(* IEC 61131-3 sources: SemaPLC/sema-plc-benchmark/spec2control-benchmark/data/st-baseline/desalination/pous/programs, 6 files *)

(* ---- main.st ---- *)
PROGRAM main
VAR
	Heartbeat : bool;
END_VAR

(* Entry point required by OpenPLC Editor v4. The process sections run as parallel program instances under task0; main only provides a scan heartbeat. *)
Heartbeat := NOT Heartbeat;

END_PROGRAM

(* ---- Section2.st ---- *)
PROGRAM Section2
VAR
	FT101_Flow_PV : real;
	FT102_Flow_PV : real;
	AT101_Analyzer_PV : real;
	AT103_Analyzer_PV : real;
	LT104_Level_PV : real;
	LT105_Level_PV : real;
	FC101_MV_Out : real;
	FC102_MV_Out : real;
	FV101_Valve_Position : real;
	FV102_Valve_Position : real;
	SP101_PctCmd : real;
	SP102_PctCmd : real;
	FlowDevAlarm101 : bool;
	FlowDevAlarm102 : bool;
	AT_101 : ANALOG_IN;
	AT_103 : ANALOG_IN;
	FC_101 : PID_BASIC;
	FC_102 : PID_BASIC;
	FT_101 : ANALOG_IN;
	FT_102 : ANALOG_IN;
	FV_101 : VALVE_ELECTRIC;
	FV_102 : VALVE_ELECTRIC;
	LT_104 : ANALOG_IN;
	LT_105 : ANALOG_IN;
	XV_102 : VALVE_ON_OFF;
	SP101_DevDelay_TON : TON;
	SP102_DevDelay_TON : TON;
	XV102NotOpen_NOT : bool;
	Contamination_OR : bool;
	FV101_Inhibit_OR : bool;
	FV102_Inhibit_OR : bool;
	SP101_PctNorm_DIV : real;
	SP101_PctScaled_MULT : real;
	SP101_PctOffset_ADD : real;
	SP101_PctToFrac_DIV : real;
	SP101_SP_EU_MULT : real;
	DL101_MULT : real;
	SP101_1p1_MULT : real;
	SP101_0p9_MULT : real;
	SP101_PV_GT_HighThresh : bool;
	SP101_PV_LT_LowThresh : bool;
	SP101_DevBand_OR : bool;
	SP102_PctNorm_DIV : real;
	SP102_PctScaled_MULT : real;
	SP102_PctOffset_ADD : real;
	SP102_PctToFrac_DIV : real;
	SP102_SP_EU_MULT : real;
	DL102_MULT : real;
	SP102_1p1_MULT : real;
	SP102_0p9_MULT : real;
	SP102_PV_GT_HighThresh : bool;
	SP102_PV_LT_LowThresh : bool;
	SP102_DevBand_OR : bool;
END_VAR

AT_101(
    PV_High := 50.0,
    Alarm_Enable := TRUE);
AT_103(
    PV_High := 35.0,
    Alarm_Enable := TRUE);
SP101_PctNorm_DIV := SP101_PctCmd / 100.0;
SP101_PctScaled_MULT := SP101_PctNorm_DIV * 59.0;
SP101_PctOffset_ADD := SP101_PctScaled_MULT + 16.0;
SP101_PctToFrac_DIV := SP101_PctOffset_ADD / 100.0;
SP101_SP_EU_MULT := SP101_PctToFrac_DIV * 5000.0;
DL101_MULT := SP101_SP_EU_MULT * 0.1;
FT_101(
    PV_High := 5500.0,
    PV_Low := 450.0,
    Scaling_Slope := 312.5,
    Scaling_Offset := -1250.0,
    Alarm_Enable := TRUE);
FC_101(
    AUTO := TRUE,
    PV := FT_101.PV,
    SP := SP101_SP_EU_MULT,
    MV_MIN := 0.0,
    MV_MAX := 100.0,
    X0 := 0.0,
    KP := 2.5,
    TR := 0.8,
    TD := 0.2,
    Deviation_Limit := DL101_MULT,
    Inhibit := FT_101.General_Fault);
SP102_PctNorm_DIV := SP102_PctCmd / 100.0;
SP102_PctScaled_MULT := SP102_PctNorm_DIV * 59.0;
SP102_PctOffset_ADD := SP102_PctScaled_MULT + 16.0;
SP102_PctToFrac_DIV := SP102_PctOffset_ADD / 100.0;
SP102_SP_EU_MULT := SP102_PctToFrac_DIV * 3000.0;
DL102_MULT := SP102_SP_EU_MULT * 0.1;
FT_102(
    PV_High := 3300.0,
    PV_Low := 270.0,
    Scaling_Slope := 187.5,
    Scaling_Offset := -750.0,
    Alarm_Enable := TRUE);
FC_102(
    AUTO := TRUE,
    PV := FT_102.PV,
    SP := SP102_SP_EU_MULT,
    MV_MIN := 0.0,
    MV_MAX := 100.0,
    X0 := 0.0,
    KP := 2.5,
    TR := 0.8,
    TD := 0.2,
    Deviation_Limit := DL102_MULT,
    Inhibit := FT_102.General_Fault);
Contamination_OR := AT_101.High_Alarm OR AT_103.High_Alarm;
LT_104(
    PV_Low := 2.0,
    Alarm_Enable := TRUE);
LT_105(
    Alarm_Enable := TRUE);
XV_102(
    Inhibit := Contamination_OR);
XV102NotOpen_NOT := NOT XV_102.FB_Opened;
FV101_Inhibit_OR := XV102NotOpen_NOT OR Contamination_OR OR LT_104.Low_Alarm OR LT_105.High_Alarm OR FT_101.General_Fault;
FV_101(
    Control_Signal := FC_101.XOUT,
    Manual_Mode := FALSE,
    Manual_Position := 0.0,
    Open_Limit := 100.0,
    Close_Limit := 0.0,
    Inhibit := FV101_Inhibit_OR);
FV102_Inhibit_OR := XV102NotOpen_NOT OR Contamination_OR OR LT_104.Low_Alarm OR LT_105.High_Alarm OR FT_102.General_Fault;
FV_102(
    Control_Signal := FC_102.XOUT,
    Manual_Mode := FALSE,
    Manual_Position := 0.0,
    Open_Limit := 100.0,
    Close_Limit := 0.0,
    Inhibit := FV102_Inhibit_OR);
SP101_1p1_MULT := SP101_SP_EU_MULT * 1.1;
SP101_PV_GT_HighThresh := (FT_101.PV > SP101_1p1_MULT);
SP101_0p9_MULT := SP101_SP_EU_MULT * 0.9;
SP101_PV_LT_LowThresh := (FT_101.PV < SP101_0p9_MULT);
SP101_DevBand_OR := SP101_PV_GT_HighThresh OR SP101_PV_LT_LowThresh;
SP101_DevDelay_TON(
    IN := SP101_DevBand_OR,
    PT := T#30s);
SP102_1p1_MULT := SP102_SP_EU_MULT * 1.1;
SP102_PV_GT_HighThresh := (FT_102.PV > SP102_1p1_MULT);
SP102_0p9_MULT := SP102_SP_EU_MULT * 0.9;
SP102_PV_LT_LowThresh := (FT_102.PV < SP102_0p9_MULT);
SP102_DevBand_OR := SP102_PV_GT_HighThresh OR SP102_PV_LT_LowThresh;
SP102_DevDelay_TON(
    IN := SP102_DevBand_OR,
    PT := T#30s);

(* Outputs published to other sections / HMI. *)
FT101_Flow_PV := FT_101.PV;
FT102_Flow_PV := FT_102.PV;
AT101_Analyzer_PV := AT_101.PV;
AT103_Analyzer_PV := AT_103.PV;
LT104_Level_PV := LT_104.PV;
LT105_Level_PV := LT_105.PV;
FC101_MV_Out := FC_101.XOUT;
FC102_MV_Out := FC_102.XOUT;
FV101_Valve_Position := FV_101.Valve_Position;
FV102_Valve_Position := FV_102.Valve_Position;
FlowDevAlarm101 := SP101_DevDelay_TON.Q;
FlowDevAlarm102 := SP102_DevDelay_TON.Q;

END_PROGRAM

(* ---- Section3.st ---- *)
PROGRAM Section3
VAR
	FT102_SP_FromRatio : real;
	FV105_Feedback_Position : real;
	FFIC_103 : RATIO_CONTROL;
	FIC_104 : PID_BASIC;
	FV_105 : VALVE_ELECTRIC;
	FT_101 : ANALOG_IN;
	FT_102 : ANALOG_IN;
	PT_103 : ANALOG_IN;
	PT_104 : ANALOG_IN;
	PIT_105 : ANALOG_IN;
	PIT_106 : ANALOG_IN;
	PT_108 : ANALOG_IN;
	SW_SCREEN_1 : BOOL_INPUT;
	SW_SCREEN_2 : BOOL_INPUT;
	SW_SCREEN_3 : BOOL_INPUT;
	SW_SCREEN_4 : BOOL_INPUT;
	SW_SCREEN_5 : BOOL_INPUT;
	SW_SCREEN_6 : BOOL_INPUT;
	RES_SCREEN_1 : BOOL_INPUT;
	RES_SCREEN_2 : BOOL_INPUT;
	RES_SCREEN_3 : BOOL_INPUT;
	RES_SCREEN_4 : BOOL_INPUT;
	LowFlowOn : bool;
	LowFlowOff : bool;
	LowFlowLatch : bool;
	AutoEnableInv : bool;
	DownstreamOutOfRange : bool;
	SupplyPressureTrip : bool;
	ValveInhibit : bool;
	Screen1Others : bool;
	Screen2Others : bool;
	Screen3Others : bool;
	Screen4Others : bool;
	Screen5Others : bool;
	Screen6Others : bool;
	Res1Others : bool;
	Res2Others : bool;
	Res3Others : bool;
	Res4Others : bool;
	Screen1WithAnother : bool;
	Screen2WithAnother : bool;
	Screen3WithAnother : bool;
	Screen4WithAnother : bool;
	Screen5WithAnother : bool;
	Screen6WithAnother : bool;
	Res1WithAnother : bool;
	Res2WithAnother : bool;
	Res3WithAnother : bool;
	Res4WithAnother : bool;
	ScreenConflict : bool;
	RatioInhibit : bool;
END_VAR

FT_101(
    PV_Low := 50.0,
    Scaling_Slope := 31.25,
    Scaling_Offset := -125.0,
    Alarm_Enable := TRUE);
FT_102(
    Scaling_Slope := 31.25,
    Scaling_Offset := -125.0);
PIT_105(
    Alarm_Enable := TRUE);
PIT_106(
    Alarm_Enable := TRUE);
DownstreamOutOfRange := PIT_105.Low_Alarm OR PIT_105.High_Alarm OR PIT_106.Low_Alarm OR PIT_106.High_Alarm;
LowFlowOff := (FT_101.PV > 50.0);
LowFlowOn := (FT_101.PV < 50.0);
LowFlowLatch := (LowFlowOn OR LowFlowLatch) AND NOT LowFlowOff;
AutoEnableInv := NOT LowFlowLatch;
FIC_104(
    AUTO := AutoEnableInv,
    PV := FT_102.PV,
    SP := FFIC_103.SlaveSP);
PT_108(
    PV_High := 9.0,
    PV_Low := 5.0,
    Alarm_Enable := TRUE);
SupplyPressureTrip := PT_108.Low_Alarm OR PT_108.High_Alarm;
ValveInhibit := DownstreamOutOfRange OR SupplyPressureTrip;
FV_105(
    Control_Signal := FIC_104.XOUT,
    Timeout := T#2s,
    Inhibit := ValveInhibit);
PT_103(
    Alarm_Enable := TRUE);
PT_104(
    Alarm_Enable := TRUE);
RES_SCREEN_1();
RES_SCREEN_2();
RES_SCREEN_3();
RES_SCREEN_4();
SW_SCREEN_1();
SW_SCREEN_2();
SW_SCREEN_3();
SW_SCREEN_4();
SW_SCREEN_5();
SW_SCREEN_6();
Res1Others := SW_SCREEN_1.Bool_Out OR SW_SCREEN_2.Bool_Out OR SW_SCREEN_3.Bool_Out OR SW_SCREEN_4.Bool_Out OR SW_SCREEN_5.Bool_Out OR SW_SCREEN_6.Bool_Out OR RES_SCREEN_2.Bool_Out OR RES_SCREEN_3.Bool_Out OR RES_SCREEN_4.Bool_Out;
Res1WithAnother := RES_SCREEN_1.Bool_Out AND Res1Others;
Res2Others := SW_SCREEN_1.Bool_Out OR SW_SCREEN_2.Bool_Out OR SW_SCREEN_3.Bool_Out OR SW_SCREEN_4.Bool_Out OR SW_SCREEN_5.Bool_Out OR SW_SCREEN_6.Bool_Out OR RES_SCREEN_1.Bool_Out OR RES_SCREEN_3.Bool_Out OR RES_SCREEN_4.Bool_Out;
Res2WithAnother := RES_SCREEN_2.Bool_Out AND Res2Others;
Res3Others := SW_SCREEN_1.Bool_Out OR SW_SCREEN_2.Bool_Out OR SW_SCREEN_3.Bool_Out OR SW_SCREEN_4.Bool_Out OR SW_SCREEN_5.Bool_Out OR SW_SCREEN_6.Bool_Out OR RES_SCREEN_1.Bool_Out OR RES_SCREEN_2.Bool_Out OR RES_SCREEN_4.Bool_Out;
Res3WithAnother := RES_SCREEN_3.Bool_Out AND Res3Others;
Res4Others := SW_SCREEN_1.Bool_Out OR SW_SCREEN_2.Bool_Out OR SW_SCREEN_3.Bool_Out OR SW_SCREEN_4.Bool_Out OR SW_SCREEN_5.Bool_Out OR SW_SCREEN_6.Bool_Out OR RES_SCREEN_1.Bool_Out OR RES_SCREEN_2.Bool_Out OR RES_SCREEN_3.Bool_Out;
Res4WithAnother := RES_SCREEN_4.Bool_Out AND Res4Others;
Screen1Others := SW_SCREEN_2.Bool_Out OR SW_SCREEN_3.Bool_Out OR SW_SCREEN_4.Bool_Out OR SW_SCREEN_5.Bool_Out OR SW_SCREEN_6.Bool_Out OR RES_SCREEN_1.Bool_Out OR RES_SCREEN_2.Bool_Out OR RES_SCREEN_3.Bool_Out OR RES_SCREEN_4.Bool_Out;
Screen1WithAnother := SW_SCREEN_1.Bool_Out AND Screen1Others;
Screen2Others := SW_SCREEN_1.Bool_Out OR SW_SCREEN_3.Bool_Out OR SW_SCREEN_4.Bool_Out OR SW_SCREEN_5.Bool_Out OR SW_SCREEN_6.Bool_Out OR RES_SCREEN_1.Bool_Out OR RES_SCREEN_2.Bool_Out OR RES_SCREEN_3.Bool_Out OR RES_SCREEN_4.Bool_Out;
Screen2WithAnother := SW_SCREEN_2.Bool_Out AND Screen2Others;
Screen3Others := SW_SCREEN_1.Bool_Out OR SW_SCREEN_2.Bool_Out OR SW_SCREEN_4.Bool_Out OR SW_SCREEN_5.Bool_Out OR SW_SCREEN_6.Bool_Out OR RES_SCREEN_1.Bool_Out OR RES_SCREEN_2.Bool_Out OR RES_SCREEN_3.Bool_Out OR RES_SCREEN_4.Bool_Out;
Screen3WithAnother := SW_SCREEN_3.Bool_Out AND Screen3Others;
Screen4Others := SW_SCREEN_1.Bool_Out OR SW_SCREEN_2.Bool_Out OR SW_SCREEN_3.Bool_Out OR SW_SCREEN_5.Bool_Out OR SW_SCREEN_6.Bool_Out OR RES_SCREEN_1.Bool_Out OR RES_SCREEN_2.Bool_Out OR RES_SCREEN_3.Bool_Out OR RES_SCREEN_4.Bool_Out;
Screen4WithAnother := SW_SCREEN_4.Bool_Out AND Screen4Others;
Screen5Others := SW_SCREEN_1.Bool_Out OR SW_SCREEN_2.Bool_Out OR SW_SCREEN_3.Bool_Out OR SW_SCREEN_4.Bool_Out OR SW_SCREEN_6.Bool_Out OR RES_SCREEN_1.Bool_Out OR RES_SCREEN_2.Bool_Out OR RES_SCREEN_3.Bool_Out OR RES_SCREEN_4.Bool_Out;
Screen5WithAnother := SW_SCREEN_5.Bool_Out AND Screen5Others;
Screen6Others := SW_SCREEN_1.Bool_Out OR SW_SCREEN_2.Bool_Out OR SW_SCREEN_3.Bool_Out OR SW_SCREEN_4.Bool_Out OR SW_SCREEN_5.Bool_Out OR RES_SCREEN_1.Bool_Out OR RES_SCREEN_2.Bool_Out OR RES_SCREEN_3.Bool_Out OR RES_SCREEN_4.Bool_Out;
Screen6WithAnother := SW_SCREEN_6.Bool_Out AND Screen6Others;
ScreenConflict := Screen1WithAnother OR Screen2WithAnother OR Screen3WithAnother OR Screen4WithAnother OR Screen5WithAnother OR Screen6WithAnother OR Res1WithAnother OR Res2WithAnother OR Res3WithAnother OR Res4WithAnother;
RatioInhibit := PT_103.Low_Alarm OR DownstreamOutOfRange OR SupplyPressureTrip OR FV_105.Position_Error OR ScreenConflict OR FIC_104.Deviation_Alarm OR LowFlowLatch OR PT_104.Low_Alarm;
FFIC_103(
    PrimaryPV := FT_101.PV,
    SecondaryPV := FT_102.PV,
    RatioSP := 2.0,
    MV_MIN := 0.0,
    MV_MAX := 500.0,
    Inhibit := RatioInhibit);

(* Outputs published to other sections / HMI. *)
FT102_SP_FromRatio := FFIC_103.SlaveSP;
FV105_Feedback_Position := FV_105.Feedback_Pos;

END_PROGRAM

(* ---- Section4.st ---- *)
PROGRAM Section4
VAR
	FT_101_Flow_PV_m3ph : real;
	LT_101_SumpLevel_m : real;
	FIC_101_MV_Percent : real;
	FIC_101_SP_m3ph : real;
	Flow_Deviation_Alarm : bool;
	FT_101 : ANALOG_IN;
	LT_101 : ANALOG_IN;
	FIC_101 : PID_BASIC;
	VFD_101A : MOTOR_VSD;
	VFD_101B : MOTOR_VSD;
	VFD_101C : MOTOR_VSD;
	VFD_101D : MOTOR_VSD;
	SPUMP_201A : MOTOR_ON_OFF;
	SPUMP_201B : MOTOR_ON_OFF;
	M103A : DIGITAL_IN;
	M103B : DIGITAL_IN;
	M103C : DIGITAL_IN;
	M103D : DIGITAL_IN;
	FlowDeviationHold : TON;
	SumpLevelOutOfRange : bool;
	Inhibit_101A : bool;
	Inhibit_101B : bool;
	Inhibit_101C : bool;
	Inhibit_101D : bool;
END_VAR

FT_101(
    Scaling_Slope := 31.25,
    Scaling_Offset := -125.0,
    Alarm_Enable := TRUE);
LT_101(
    PV_High := 9.0,
    PV_Low := 1.5,
    Scaling_Slope := 0.625,
    Scaling_Offset := -2.5,
    Alarm_Enable := TRUE);
SumpLevelOutOfRange := LT_101.Low_Alarm OR LT_101.High_Alarm;
FIC_101(
    AUTO := TRUE,
    PV := FT_101.PV,
    SP := FIC_101_SP_m3ph,
    MV_MIN := 0.0,
    MV_MAX := 100.0,
    X0 := 0.0,
    KP := 2.5,
    TR := 0.8,
    TD := 0.2,
    Deviation_Limit := 10.0,
    Inhibit := SumpLevelOutOfRange);
M103A();
Inhibit_101A := SumpLevelOutOfRange OR M103A.DI_Out OR VFD_101A.FB_Fault;
VFD_101A(
    Speed_SP := FIC_101.XOUT,
    Inhibit := Inhibit_101A);
M103B();
Inhibit_101B := SumpLevelOutOfRange OR M103B.DI_Out OR VFD_101B.FB_Fault;
VFD_101B(
    Inhibit := Inhibit_101B);
M103C();
Inhibit_101C := SumpLevelOutOfRange OR M103C.DI_Out OR VFD_101C.FB_Fault;
VFD_101C(
    Inhibit := Inhibit_101C);
M103D();
Inhibit_101D := SumpLevelOutOfRange OR M103D.DI_Out OR VFD_101D.FB_Fault;
VFD_101D(
    Inhibit := Inhibit_101D);
SPUMP_201A();
SPUMP_201B();
FlowDeviationHold(
    IN := FIC_101.Deviation_Alarm,
    PT := T#30s);

(* Outputs published to other sections / HMI. *)
Flow_Deviation_Alarm := FlowDeviationHold.Q;
FT_101_Flow_PV_m3ph := FT_101.PV;
LT_101_SumpLevel_m := LT_101.PV;
FIC_101_MV_Percent := FIC_101.XOUT;

END_PROGRAM

(* ---- Section5.st ---- *)
PROGRAM Section5
VAR
	FT_301_FlowRate_PV : real;
	LT_301_Level_PV : real;
	FIC_301_MV_FlowControl_Percent : real;
	XV_107_Open_FB : bool;
	FT_301 : ANALOG_IN;
	LT_301 : ANALOG_IN;
	FIC_301 : PID_BASIC;
	FV_301 : VALVE_ELECTRIC;
	XV_107 : VALVE_ON_OFF;
	UMP_301A : MOTOR_VSD;
	UMP_301B : MOTOR_VSD;
	ANK_301 : BOOL_INPUT;
	PAH_103 : DIGITAL_IN;
	TAH_101 : DIGITAL_IN;
	NotXVOpen_NOT : bool;
	PumpsAvailable_OR : bool;
	NotPumpsAvailable_NOT : bool;
	LevelNotAbove20_NOT : bool;
	PumpInhibit_OR : bool;
	ValveTrips_OR : bool;
	PIDInhibit_OR : bool;
END_VAR

FT_301(
    PV_High := 48.0,
    PV_Low := 8.0,
    Scaling_Slope := 3.125,
    Scaling_Offset := -12.5,
    Alarm_Enable := TRUE);
LT_301(
    Alarm_Enable := TRUE);
ANK_301();
LevelNotAbove20_NOT := NOT LT_301.High_Alarm;
UMP_301A(
    Speed_SP := FIC_301.XOUT,
    Inhibit := PumpInhibit_OR);
UMP_301B(
    Inhibit := PumpInhibit_OR);
PumpsAvailable_OR := UMP_301A.FB_Ready OR UMP_301B.FB_Ready;
NotPumpsAvailable_NOT := NOT PumpsAvailable_OR;
XV_107();
NotXVOpen_NOT := NOT XV_107.FB_Opened;
PumpInhibit_OR := NotXVOpen_NOT OR NotPumpsAvailable_NOT OR ANK_301.Bool_Out OR LT_301.Low_Alarm OR LevelNotAbove20_NOT;
PAH_103();
TAH_101();
ValveTrips_OR := PAH_103.DI_Out OR TAH_101.DI_Out OR LT_301.Low_Alarm OR ANK_301.Bool_Out;
PIDInhibit_OR := PumpInhibit_OR OR ValveTrips_OR;
FIC_301(
    PV := FT_301.PV,
    SP := 30.0,
    MV_MIN := 5.0,
    MV_MAX := 95.0,
    X0 := UMP_301A.FB_ActualSpeed,
    KP := 1.8,
    TR := 0.5,
    TD := 0.05,
    Inhibit := PIDInhibit_OR);
FV_301(
    Open_Limit := 100.0,
    Close_Limit := 0.0,
    Inhibit := ValveTrips_OR);

(* Outputs published to other sections / HMI. *)
FT_301_FlowRate_PV := FT_301.PV;
LT_301_Level_PV := LT_301.PV;
FIC_301_MV_FlowControl_Percent := FIC_301.XOUT;
XV_107_Open_FB := XV_107.FB_Opened;

END_PROGRAM

(* ---- Section6.st ---- *)
PROGRAM Section6
VAR
	FIT101_BypassFlow_PV : real;
	FIT102_SamplingFlow_PV : real;
	FIC104_SamplingFlow_SP : real;
	FIC104_ActiveRatio : real;
	AT105_Permissive : bool;
	LV103_Permissive : bool;
	FIT_101 : ANALOG_IN;
	FIT_102 : ANALOG_IN;
	FIC_104 : RATIO_CONTROL;
	FIC_104_SLAVE : PID_BASIC;
	FV_102 : VALVE_ELECTRIC;
	AT_105 : BOOL_INPUT;
	MasterInhibit_OR : bool;
	LV103_Permissive_NOT : bool;
END_VAR

FIT_101(
    Scaling_Slope := 62.5,
    Scaling_Offset := -250.0,
    Alarm_Enable := TRUE);
FIT_102(
    Alarm_Enable := TRUE);
AT_105(
    Bool_In := AT105_Permissive,
    Alarm_OnTrue := FALSE,
    Alarm_OnFalse := TRUE,
    Latch_Enable := TRUE);
LV103_Permissive_NOT := NOT LV103_Permissive;
MasterInhibit_OR := FIT_101.Low_Alarm OR FIT_101.General_Fault OR AT_105.Alarm_Active OR LV103_Permissive_NOT;
FIC_104(
    Auto := TRUE,
    PrimaryPV := FIT_101.PV,
    SecondaryPV := FIT_102.PV,
    RatioSP := 0.1,
    MV_MIN := 0.0,
    MV_MAX := 200.0,
    Inhibit := MasterInhibit_OR);
FIC_104_SLAVE(
    AUTO := TRUE,
    PV := FIT_102.PV,
    SP := FIC_104.SlaveSP,
    MV_MIN := 0.0,
    MV_MAX := 100.0,
    X0 := 0.0,
    KP := 1.0,
    TR := 10.0,
    TD := 0.0,
    Deviation_Limit := 20.0,
    Inhibit := MasterInhibit_OR);
FV_102(
    Control_Signal := FIC_104_SLAVE.XOUT,
    Manual_Mode := FALSE,
    Open_Limit := 100.0,
    Close_Limit := 0.0,
    Inhibit := MasterInhibit_OR);

(* Outputs published to other sections / HMI. *)
FIT101_BypassFlow_PV := FIT_101.PV;
FIT102_SamplingFlow_PV := FIT_102.PV;
FIC104_SamplingFlow_SP := FIC_104.SlaveSP;
FIC104_ActiveRatio := FIC_104.ActiveRatio;

END_PROGRAM
